Fanuc KAREL source: kf00114.compact.KL

PROGRAM KF00114
%STACKSIZE=65535
%PRIORITY=65535
%NOLOCKGROUP
VAR
I : INTEGER
J : INTEGER
X : REAL
Y : REAL
B : BOOLEAN
C : BOOLEAN
TXT : STRING[80]
TXT2 : STRING[80]
AI : ARRAY[4] OF INTEGER
BI : ARRAY[4] OF INTEGER
P : XYZWPR
JP : JOINTPOS9
PF : POSITION
V1 : VECTOR
V2 : VECTOR
STATUS : INTEGER
ROUTINE PADD(P1 : INTEGER) FROM KF00114
ROUTINE PADD
BEGIN
I=(P1 + 1)
END PADD
BEGIN
PADD(I)
END KF00114
